SUBAPPLICATION Uebung_254b_AX (* PWM sprungartig mit Tastern: I6 = 0, I7 = 4000, I8 = 8000 auf PWM Q1, RAMP T#0ms *)
  (* Standard: 61499-2; Description: Copyright (c) 2026 Meisterschulen am Ostbahnhof This program and the accompanying materials are made available under the terms of the Eclipse Public License 2.0 which is available at https://www.eclipse.org/legal/epl-2.0/ SPDX-License-Identifier: EPL-2.0 *)
  (* Version 1.0, 2026-11-06, Franz Höpfinger, Meisterschulen am Ostbahnhof, initial API and implementation and/or initial documentation *)
  PACKAGE Uebungen;
  IMPORT logiBUS::io::DI::logiBUS_DI::Input_I6;
  IMPORT logiBUS::io::DI::logiBUS_DI::Input_I7;
  IMPORT logiBUS::io::DI::logiBUS_DI::Input_I8;
  IMPORT logiBUS::io::DI::logiBUS_DI_Events::BUTTON_PRESS_DOWN;
  IMPORT logiBUS::io::DQ::logiBUS_DO::Output_Q1;
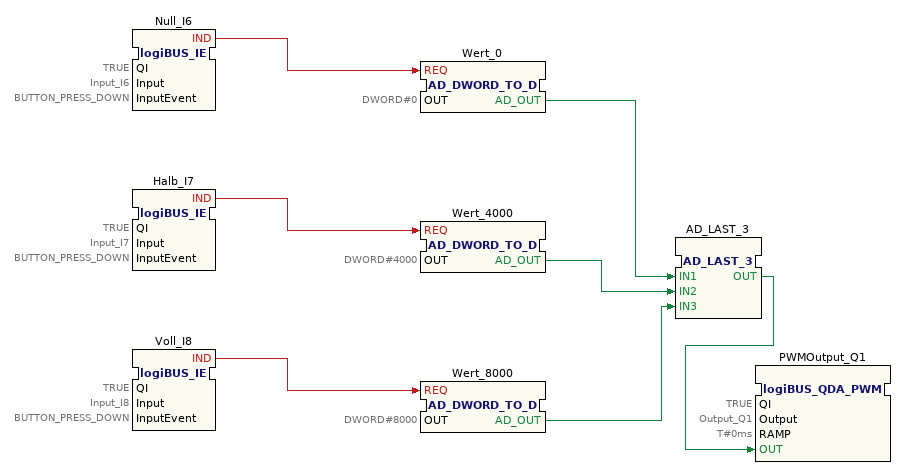
  FBS
    Null_I6 : logiBUS::io::DI::logiBUS_IE(QI := TRUE, Input := Input_I6, InputEvent := BUTTON_PRESS_DOWN);
    Wert_0 : adapter::conversion::unidirectional::AD_DWORD_TO_D(OUT := DWORD#0);
    Halb_I7 : logiBUS::io::DI::logiBUS_IE(QI := TRUE, Input := Input_I7, InputEvent := BUTTON_PRESS_DOWN);
    Wert_4000 : adapter::conversion::unidirectional::AD_DWORD_TO_D(OUT := DWORD#4000);
    Voll_I8 : logiBUS::io::DI::logiBUS_IE(QI := TRUE, Input := Input_I8, InputEvent := BUTTON_PRESS_DOWN);
    Wert_8000 : adapter::conversion::unidirectional::AD_DWORD_TO_D(OUT := DWORD#8000);
    AD_LAST_3 : adapter::events::unidirectional::AD_LAST_3;
    PWMOutput_Q1 : logiBUS::io::DQ::logiBUS_QDA_PWM(QI := TRUE, Output := Output_Q1, RAMP := T#0ms);
  END_FBS
  EVENT_CONNECTIONS
    Null_I6.IND TO Wert_0.REQ;
    Halb_I7.IND TO Wert_4000.REQ;
    Voll_I8.IND TO Wert_8000.REQ;
  END_CONNECTIONS
  ADAPTER_CONNECTIONS
    Wert_0.AD_OUT TO AD_LAST_3.IN1;
    Wert_4000.AD_OUT TO AD_LAST_3.IN2;
    Wert_8000.AD_OUT TO AD_LAST_3.IN3;
    AD_LAST_3.OUT TO PWMOutput_Q1.OUT;
  END_CONNECTIONS
END_SUBAPPLICATION
